Universal Robots PolyScope program: polyscope.in.memory.program.urp

Program <unnamed> (installation=default directory=/programs createdIn=5.21.1 lastSavedIn=5.21.1 robotSerialNumber=20255500273)
InitVariablesNode
Robot Program (runOnlyOnce=false)
  Placeholder
